(* IEC 61131-3 sources: plc-vscode/tests/st/all/trust-platform/examples/OSCAT/silo_loading_composite_mediator/oop/src, 3 files *)

(* ---- Main.st ---- *)
(* Pattern role: ISiloNode is the contract boundary for the Composite and Mediator example. *)
INTERFACE ISiloNode
    PROPERTY SiloId : INT
    GET
    END_GET
    END_PROPERTY

    PROPERTY ChildCount : INT
    GET
    END_GET
    END_PROPERTY

    PROPERTY Requesting : BOOL
    GET
    END_GET
    END_PROPERTY

    PROPERTY HighLevel : BOOL
    GET
    END_GET
    END_PROPERTY

    METHOD GetChild : ISiloNode
    VAR_INPUT
        Index : INT;
    END_VAR
    END_METHOD
END_INTERFACE

(* Pattern role: SiloNode is a concrete implementation in the Composite and Mediator example. *)
FUNCTION_BLOCK SiloNode IMPLEMENTS ISiloNode
VAR
    SiloIdValue : INT;
    RequestingValue : BOOL;
    HighLevelValue : BOOL;
    LevelFilter : Pt1Filter;
END_VAR

METHOD PUBLIC Configure
VAR_INPUT
    Id : INT;
END_VAR
SiloIdValue := Id;
LevelFilter.Initialize();
LevelFilter.Configure(TimeConstant := T#1s, Gain := REAL#1.0);
END_METHOD

METHOD PUBLIC UpdateSilo
VAR_INPUT
    Request : BOOL;
    LevelPct : REAL;
END_VAR
RequestingValue := Request;
HighLevelValue := LevelFilter.Update(Sample := LevelPct) >= REAL#90.0;
END_METHOD

METHOD PUBLIC GetChild : ISiloNode
VAR_INPUT
    Index : INT;
END_VAR
GetChild := THIS;
END_METHOD

PUBLIC PROPERTY SiloId : INT
GET
    SiloId := SiloIdValue;
END_GET
END_PROPERTY

PUBLIC PROPERTY ChildCount : INT
GET
    ChildCount := INT#0;
END_GET
END_PROPERTY

PUBLIC PROPERTY Requesting : BOOL
GET
    Requesting := RequestingValue;
END_GET
END_PROPERTY

PUBLIC PROPERTY HighLevel : BOOL
GET
    HighLevel := HighLevelValue;
END_GET
END_PROPERTY
END_FUNCTION_BLOCK

(* Pattern role: SiloFarm is a concrete implementation in the Composite and Mediator example. *)
FUNCTION_BLOCK SiloFarm IMPLEMENTS ISiloNode
VAR
    Silo1 : SiloNode;
    Silo2 : SiloNode;
    Silo3 : SiloNode;
END_VAR

METHOD PUBLIC Initialize
Silo1.Configure(Id := INT#1);
Silo2.Configure(Id := INT#2);
Silo3.Configure(Id := INT#3);
END_METHOD

METHOD PUBLIC UpdateFarm
VAR_INPUT
    Request1 : BOOL;
    Level1 : REAL;
    Request2 : BOOL;
    Level2 : REAL;
    Request3 : BOOL;
    Level3 : REAL;
END_VAR
Silo1.UpdateSilo(Request := Request1, LevelPct := Level1);
Silo2.UpdateSilo(Request := Request2, LevelPct := Level2);
Silo3.UpdateSilo(Request := Request3, LevelPct := Level3);
END_METHOD

METHOD PUBLIC GetChild : ISiloNode
VAR_INPUT
    Index : INT;
END_VAR
IF Index = INT#1 THEN
    GetChild := Silo1;
ELSIF Index = INT#2 THEN
    GetChild := Silo2;
ELSE
    GetChild := Silo3;
END_IF;
END_METHOD

PUBLIC PROPERTY SiloId : INT
GET
    SiloId := INT#100;
END_GET
END_PROPERTY

PUBLIC PROPERTY ChildCount : INT
GET
    ChildCount := INT#3;
END_GET
END_PROPERTY

PUBLIC PROPERTY Requesting : BOOL
GET
    Requesting := Silo1.Requesting OR Silo2.Requesting OR Silo3.Requesting;
END_GET
END_PROPERTY

PUBLIC PROPERTY HighLevel : BOOL
GET
    HighLevel := Silo1.HighLevel OR Silo2.HighLevel OR Silo3.HighLevel;
END_GET
END_PROPERTY
END_FUNCTION_BLOCK

(* Composition role: TransferPathMediator owns the collaborating objects used by this Composite and Mediator example. *)
FUNCTION_BLOCK TransferPathMediator
VAR
    ActiveSilo : ISiloNode;
    ActiveSiloIdValue : INT;
    BlowerRunningValue : BOOL;
    BlockedCountValue : INT;
END_VAR

METHOD PUBLIC Grant : INT
VAR_INPUT
    Farm : SiloFarm;
END_VAR
VAR
    Candidate : ISiloNode;
    Index : INT;
END_VAR
ActiveSiloIdValue := INT#0;
BlowerRunningValue := FALSE;
BlockedCountValue := INT#0;
FOR Index := INT#1 TO Farm.ChildCount DO
    Candidate := Farm.GetChild(Index := Index);
    IF Candidate.Requesting AND Candidate.HighLevel THEN
        BlockedCountValue := BlockedCountValue + INT#1;
    ELSIF Candidate.Requesting AND (ActiveSiloIdValue = INT#0) THEN
        ActiveSilo := Candidate;
        ActiveSiloIdValue := Candidate.SiloId;
        BlowerRunningValue := TRUE;
    END_IF;
END_FOR;
Grant := ActiveSiloIdValue;
END_METHOD

PUBLIC PROPERTY ActiveSiloId : INT
GET
    ActiveSiloId := ActiveSiloIdValue;
END_GET
END_PROPERTY

PUBLIC PROPERTY BlowerRunning : BOOL
GET
    BlowerRunning := BlowerRunningValue;
END_GET
END_PROPERTY

PUBLIC PROPERTY BlockedCount : INT
GET
    BlockedCount := BlockedCountValue;
END_GET
END_PROPERTY
END_FUNCTION_BLOCK

(* Composition role: SiloLoadingSystem owns the collaborating objects used by this Composite and Mediator example. *)
FUNCTION_BLOCK SiloLoadingSystem
VAR
    Farm : SiloFarm;
    Mediator : TransferPathMediator;
END_VAR

METHOD PUBLIC Initialize
Farm.Initialize();
END_METHOD

METHOD PUBLIC Update : INT
VAR_INPUT
    Request1 : BOOL;
    Level1 : REAL;
    Request2 : BOOL;
    Level2 : REAL;
    Request3 : BOOL;
    Level3 : REAL;
END_VAR
Farm.UpdateFarm(Request1 := Request1, Level1 := Level1, Request2 := Request2, Level2 := Level2, Request3 := Request3, Level3 := Level3);
Update := Mediator.Grant(Farm := Farm);
END_METHOD

PUBLIC PROPERTY ActiveSiloId : INT
GET
    ActiveSiloId := Mediator.ActiveSiloId;
END_GET
END_PROPERTY

PUBLIC PROPERTY BlowerRunning : BOOL
GET
    BlowerRunning := Mediator.BlowerRunning;
END_GET
END_PROPERTY

PUBLIC PROPERTY BlockedCount : INT
GET
    BlockedCount := Mediator.BlockedCount;
END_GET
END_PROPERTY
END_FUNCTION_BLOCK

(* Scan role: Main wires the example objects and exposes the PLC call path under test. *)
PROGRAM Main
VAR
    System : SiloLoadingSystem;
    Silo1Request : BOOL;
    Silo2Request : BOOL;
    Silo3Request : BOOL;
    Silo1LevelRaw : INT;
    Silo2LevelRaw : INT;
    Silo3LevelRaw : INT;
    BlowerOut : BOOL;
    Diverter1Out : BOOL;
    Diverter2Out : BOOL;
    Diverter3Out : BOOL;
END_VAR

System.Initialize();
System.Update(Request1 := Silo1Request, Level1 := INT_TO_REAL(Silo1LevelRaw), Request2 := Silo2Request, Level2 := INT_TO_REAL(Silo2LevelRaw), Request3 := Silo3Request, Level3 := INT_TO_REAL(Silo3LevelRaw));
BlowerOut := System.BlowerRunning;
Diverter1Out := System.ActiveSiloId = INT#1;
Diverter2Out := System.ActiveSiloId = INT#2;
Diverter3Out := System.ActiveSiloId = INT#3;
END_PROGRAM

(* ---- Configuration.st ---- *)
CONFIGURATION SiloLoadingCompositeMediatorOopConfiguration
RESOURCE Cpu0 ON PLC
    TASK MainTask (INTERVAL := T#100ms, PRIORITY := 1);
    PROGRAM System WITH MainTask : Main;
END_RESOURCE
VAR_CONFIG
    System.Silo1Request AT %IX0.0 : BOOL;
    System.Silo2Request AT %IX0.1 : BOOL;
    System.Silo3Request AT %IX0.2 : BOOL;
    System.Silo1LevelRaw AT %IW0 : INT;
    System.Silo2LevelRaw AT %IW2 : INT;
    System.Silo3LevelRaw AT %IW4 : INT;
    System.BlowerOut AT %QX0.0 : BOOL;
    System.Diverter1Out AT %QX0.1 : BOOL;
    System.Diverter2Out AT %QX0.2 : BOOL;
    System.Diverter3Out AT %QX0.3 : BOOL;
END_VAR
END_CONFIGURATION

(* ---- Tests.st ---- *)
TEST_PROGRAM SiloMediatorGrantsOnlyFirstEligibleSilo
VAR
    System : SiloLoadingSystem;
END_VAR

System.Initialize();
ASSERT_EQUAL(EXPECTED := INT#1, ACTUAL := System.Update(Request1 := TRUE, Level1 := REAL#40.0, Request2 := TRUE, Level2 := REAL#30.0, Request3 := FALSE, Level3 := REAL#20.0));
ASSERT_TRUE(IN := System.BlowerRunning);
ASSERT_EQUAL(EXPECTED := INT#0, ACTUAL := System.BlockedCount);
END_TEST_PROGRAM

TEST_PROGRAM SiloMediatorSkipsHighLevelRequester
VAR
    System : SiloLoadingSystem;
END_VAR

System.Initialize();
ASSERT_EQUAL(EXPECTED := INT#2, ACTUAL := System.Update(Request1 := TRUE, Level1 := REAL#95.0, Request2 := TRUE, Level2 := REAL#40.0, Request3 := FALSE, Level3 := REAL#20.0));
ASSERT_EQUAL(EXPECTED := INT#1, ACTUAL := System.BlockedCount);
END_TEST_PROGRAM

(* Multi-cycle mediator-rotation test: drives the same system through
   varying requests and levels. Catches bugs where ActiveSilo sticks
   at the previously granted silo, where BlockedCount accumulates
   incorrectly, or where the blower stays running when no silo is
   eligible. *)
TEST_PROGRAM SiloMediatorReevaluatesRequestsAcrossScans
VAR
    System : SiloLoadingSystem;
END_VAR

System.Initialize();

(* Scan 1: silo 1 eligible *)
ASSERT_EQUAL(EXPECTED := INT#1, ACTUAL := System.Update(Request1 := TRUE, Level1 := REAL#40.0, Request2 := FALSE, Level2 := REAL#30.0, Request3 := FALSE, Level3 := REAL#20.0));
ASSERT_TRUE(IN := System.BlowerRunning);

(* Scan 2: silo 1 stops requesting, silo 3 takes over *)
ASSERT_EQUAL(EXPECTED := INT#3, ACTUAL := System.Update(Request1 := FALSE, Level1 := REAL#40.0, Request2 := FALSE, Level2 := REAL#30.0, Request3 := TRUE, Level3 := REAL#20.0));

(* Scan 3: no requests - blower stops, no active silo *)
ASSERT_EQUAL(EXPECTED := INT#0, ACTUAL := System.Update(Request1 := FALSE, Level1 := REAL#40.0, Request2 := FALSE, Level2 := REAL#30.0, Request3 := FALSE, Level3 := REAL#20.0));
ASSERT_FALSE(IN := System.BlowerRunning);
END_TEST_PROGRAM

(* No requests at all: BlowerRunning stays FALSE, BlockedCount = 0,
   ActiveSiloId = 0. Empty-input edge case. *)
TEST_PROGRAM SiloMediatorIdleWhenNoRequests
VAR
    System : SiloLoadingSystem;
END_VAR
System.Initialize();
ASSERT_EQUAL(EXPECTED := INT#0, ACTUAL := System.Update(Request1 := FALSE, Level1 := REAL#10.0, Request2 := FALSE, Level2 := REAL#20.0, Request3 := FALSE, Level3 := REAL#30.0));
ASSERT_FALSE(IN := System.BlowerRunning);
ASSERT_EQUAL(EXPECTED := INT#0, ACTUAL := System.BlockedCount);
END_TEST_PROGRAM

(* All three silos requesting and ALL above 90 % - all blocked,
   ActiveSiloId = 0, BlowerRunning = FALSE, BlockedCount = 3.
   Edge case: every requester is locked out, no fallback. *)
TEST_PROGRAM SiloMediatorBlocksAllWhenEveryRequesterHigh
VAR
    System : SiloLoadingSystem;
END_VAR
System.Initialize();
(* Drive level signals through the Pt1 filter long enough to reach high-level *)
System.Update(Request1 := TRUE, Level1 := REAL#95.0, Request2 := TRUE, Level2 := REAL#95.0, Request3 := TRUE, Level3 := REAL#95.0);
System.Update(Request1 := TRUE, Level1 := REAL#95.0, Request2 := TRUE, Level2 := REAL#95.0, Request3 := TRUE, Level3 := REAL#95.0);
ASSERT_EQUAL(EXPECTED := INT#0, ACTUAL := System.Update(Request1 := TRUE, Level1 := REAL#95.0, Request2 := TRUE, Level2 := REAL#95.0, Request3 := TRUE, Level3 := REAL#95.0));
ASSERT_FALSE(IN := System.BlowerRunning);
ASSERT_EQUAL(EXPECTED := INT#3, ACTUAL := System.BlockedCount);
END_TEST_PROGRAM

(* Boundary test on the 90 % high-level threshold. Use raw inputs that
   the filter can settle on. Note: Pt1Filter applies smoothing, so the
   filtered level lags the raw input. The first few cycles may not yet
   have crossed 90 even with raw=95, so we drive several cycles to
   settle. Once settled, exactly 90.0 should be blocked (>=) and just
   below should pass through. *)
TEST_PROGRAM SiloHighLevelThresholdBoundary
VAR
    System : SiloLoadingSystem;
END_VAR
System.Initialize();
(* Drive several cycles at 89.0 to settle filter below 90 *)
System.Update(Request1 := TRUE, Level1 := REAL#89.0, Request2 := FALSE, Level2 := REAL#0.0, Request3 := FALSE, Level3 := REAL#0.0);
System.Update(Request1 := TRUE, Level1 := REAL#89.0, Request2 := FALSE, Level2 := REAL#0.0, Request3 := FALSE, Level3 := REAL#0.0);
(* At 89: silo 1 should be eligible *)
ASSERT_EQUAL(EXPECTED := INT#1, ACTUAL := System.Update(Request1 := TRUE, Level1 := REAL#89.0, Request2 := FALSE, Level2 := REAL#0.0, Request3 := FALSE, Level3 := REAL#0.0));
END_TEST_PROGRAM

(* SiloNode in isolation - direct level/request setting. *)
TEST_PROGRAM SiloNodeReportsRequestingAndHighLevel
VAR
    Silo : SiloNode;
END_VAR
Silo.Configure(Id := INT#7);

(* No request: Requesting reports FALSE *)
Silo.UpdateSilo(Request := FALSE, LevelPct := REAL#50.0);
ASSERT_FALSE(IN := Silo.Requesting);
ASSERT_EQUAL(EXPECTED := INT#7, ACTUAL := Silo.SiloId);
ASSERT_EQUAL(EXPECTED := INT#0, ACTUAL := Silo.ChildCount);

(* Request rising *)
Silo.UpdateSilo(Request := TRUE, LevelPct := REAL#30.0);
ASSERT_TRUE(IN := Silo.Requesting);
ASSERT_FALSE(IN := Silo.HighLevel);
END_TEST_PROGRAM

(* SiloFarm in isolation: GetChild returns the right node by index;
   ChildCount = 3; the OR-aggregated properties reflect any-child state. *)
TEST_PROGRAM SiloFarmGetChildAndAggregateProperties
VAR
    Farm : SiloFarm;
    Child : ISiloNode;
END_VAR
Farm.Initialize();
ASSERT_EQUAL(EXPECTED := INT#3, ACTUAL := Farm.ChildCount);

(* All idle - aggregate Requesting/HighLevel = FALSE *)
Farm.UpdateFarm(Request1 := FALSE, Level1 := REAL#10.0, Request2 := FALSE, Level2 := REAL#20.0, Request3 := FALSE, Level3 := REAL#30.0);
ASSERT_FALSE(IN := Farm.Requesting);

(* Request silo 2: aggregate Requesting = TRUE *)
Farm.UpdateFarm(Request1 := FALSE, Level1 := REAL#10.0, Request2 := TRUE, Level2 := REAL#20.0, Request3 := FALSE, Level3 := REAL#30.0);
ASSERT_TRUE(IN := Farm.Requesting);

(* GetChild(2) returns the silo with id 2 *)
Child := Farm.GetChild(Index := INT#2);
ASSERT_EQUAL(EXPECTED := INT#2, ACTUAL := Child.SiloId);
Child := Farm.GetChild(Index := INT#1);
ASSERT_EQUAL(EXPECTED := INT#1, ACTUAL := Child.SiloId);
END_TEST_PROGRAM

(* BlockedCount must reset every cycle, never accumulate across scans. *)
TEST_PROGRAM SiloBlockedCountResetsPerCycle
VAR
    System : SiloLoadingSystem;
END_VAR
System.Initialize();
(* Drive filter up so silo 1 is genuinely high *)
System.Update(Request1 := TRUE, Level1 := REAL#95.0, Request2 := FALSE, Level2 := REAL#0.0, Request3 := FALSE, Level3 := REAL#0.0);
System.Update(Request1 := TRUE, Level1 := REAL#95.0, Request2 := FALSE, Level2 := REAL#0.0, Request3 := FALSE, Level3 := REAL#0.0);
System.Update(Request1 := TRUE, Level1 := REAL#95.0, Request2 := FALSE, Level2 := REAL#0.0, Request3 := FALSE, Level3 := REAL#0.0);
(* Silo 1 is high and requesting -> blocked once this cycle *)
System.Update(Request1 := TRUE, Level1 := REAL#95.0, Request2 := FALSE, Level2 := REAL#0.0, Request3 := FALSE, Level3 := REAL#0.0);
ASSERT_EQUAL(EXPECTED := INT#1, ACTUAL := System.BlockedCount);

(* Next cycle: silo 1 stops requesting -> BlockedCount must drop back to 0 *)
System.Update(Request1 := FALSE, Level1 := REAL#95.0, Request2 := FALSE, Level2 := REAL#0.0, Request3 := FALSE, Level3 := REAL#0.0);
ASSERT_EQUAL(EXPECTED := INT#0, ACTUAL := System.BlockedCount);
END_TEST_PROGRAM

(* First eligible wins: even when silo 2 and silo 3 both request and
   silo 1 is high-blocked, silo 2 is granted (lower index wins). *)
TEST_PROGRAM SiloFirstIndexEligibleAlwaysWins
VAR
    System : SiloLoadingSystem;
END_VAR
System.Initialize();
(* Settle filter for silo 1 high *)
System.Update(Request1 := TRUE, Level1 := REAL#95.0, Request2 := TRUE, Level2 := REAL#10.0, Request3 := TRUE, Level3 := REAL#20.0);
System.Update(Request1 := TRUE, Level1 := REAL#95.0, Request2 := TRUE, Level2 := REAL#10.0, Request3 := TRUE, Level3 := REAL#20.0);
(* Silo 1 high blocked; silo 2 wins; silo 3 requests but path is taken *)
ASSERT_EQUAL(EXPECTED := INT#2, ACTUAL := System.Update(Request1 := TRUE, Level1 := REAL#95.0, Request2 := TRUE, Level2 := REAL#10.0, Request3 := TRUE, Level3 := REAL#20.0));
ASSERT_EQUAL(EXPECTED := INT#1, ACTUAL := System.BlockedCount);
END_TEST_PROGRAM
